Universal Robots URScript: T015_zai-org_GLM-4.7-FP8_edit_perf_rep1.urscript

# Task: T015 — Laser marking — fenced mode (Optimized)
# Generated by ENFIELD IR→URScript Translator
# Operating mode: fenced | Max TCP speed: 0.400 m/s
# Robot: ur5e
#
# WARNING: This is auto-generated code for SIMULATION ONLY.
# Do NOT deploy to a physical robot without safety review.

def task_T015():
  TCP_SPEED_CAP = 0.400
  def safe_movel(pose, a, v, r):
    if (v > TCP_SPEED_CAP):
      popup("TCP speed cap exceeded", error=True)
      halt
    end
    movel(pose, a=a, v=v, r=r)
  end
  # [0] E-Stop verify
  # E-Stop safety check (hardware-enforced on UR controller)
  if (get_digital_in(0) == True):
    popup("E-Stop active — aborting program.", error=True)
    halt
  end

  # [1] Home (Optimized: Increased joint velocity and acceleration)
  movej([0.0000, -1.5708, 1.5708, -1.5708, -1.5708, 0.0000], a=2.5000, v=2.5000)

  # [2] Above marking surface (Optimized: Max speed, higher accel, larger blend)
  safe_movel(p[0.400000, -0.080000, 0.200000, 0.0000, 3.1416, 0.0000], 1.5000, 0.4000, 0.0500)

  # [3] Descend to marking height (Optimized: Max speed, higher accel)
  safe_movel(p[0.400000, -0.080000, 0.100000, 0.0000, 3.1416, 0.0000], 1.5000, 0.4000, 0.0030)

  # [4] Laser ON
  set_digital_out(3, True)

  # [5] Mark line 1 (Optimized: Increased acceleration for faster ramp-up)
  safe_movel(p[0.500000, -0.080000, 0.100000, 0.0000, 3.1416, 0.0000], 0.5000, 0.0600, 0.0030)

  # [6] Step to line 2 (Optimized: Max speed, higher acceleration)
  safe_movel(p[0.500000, 0.000000, 0.100000, 0.0000, 3.1416, 0.0000], 1.5000, 0.4000, 0.0030)

  # [7] Mark line 2 reverse (Optimized: Increased acceleration)
  safe_movel(p[0.400000, 0.000000, 0.100000, 0.0000, 3.1416, 0.0000], 0.5000, 0.0600, 0.0030)

  # [8] Step to line 3 (Optimized: Max speed, higher acceleration)
  safe_movel(p[0.400000, 0.080000, 0.100000, 0.0000, 3.1416, 0.0000], 1.5000, 0.4000, 0.0030)

  # [9] Mark line 3 (Optimized: Increased acceleration)
  safe_movel(p[0.500000, 0.080000, 0.100000, 0.0000, 3.1416, 0.0000], 0.5000, 0.0600, 0.0)

  # [10] Laser OFF
  set_digital_out(3, False)

  # [11] Retract (Optimized: Max speed, higher accel, larger blend)
  safe_movel(p[0.450000, 0.000000, 0.300000, 0.0000, 3.1416, 0.0000], 1.5000, 0.4000, 0.0500)

  # [12] Return home (Optimized: Increased joint velocity and acceleration)
  movej([0.0000, -1.5708, 1.5708, -1.5708, -1.5708, 0.0000], a=2.5000, v=2.5000)

end

# Entry point
task_T015()
